// Jugement d'un résultat (docs/04 § 5)
{attribute 'qualified_only'}
{attribute 'strict'}
TYPE E_Judgement :
(
    None := 0,
    Ok := 1,
    Nok := 2,
    High := 3,
    Low := 4
) USINT;
END_TYPE

(* stored: Version 1.1.0.1, ProductVersion 3.1.4024.12
   DUT E_Judgement: Id {58f5ec62-4990-5269-96ef-79c711bd3892} *)
